{attribute 'qualified_only'}
VAR_GLOBAL CONSTANT
	JSON_DOCUMENT_CHAR_SIZE : UINT := 25000;
	ERROR_MESSAGE_WIDE_CHAR_SIZE : UINT := 500;
END_VAR

(* stored: Version 1.1.0.1
   GVL Parameters: Id {60b8aa99-fae2-4f0a-ac60-38ea97572fc5}, ParameterList True *)
